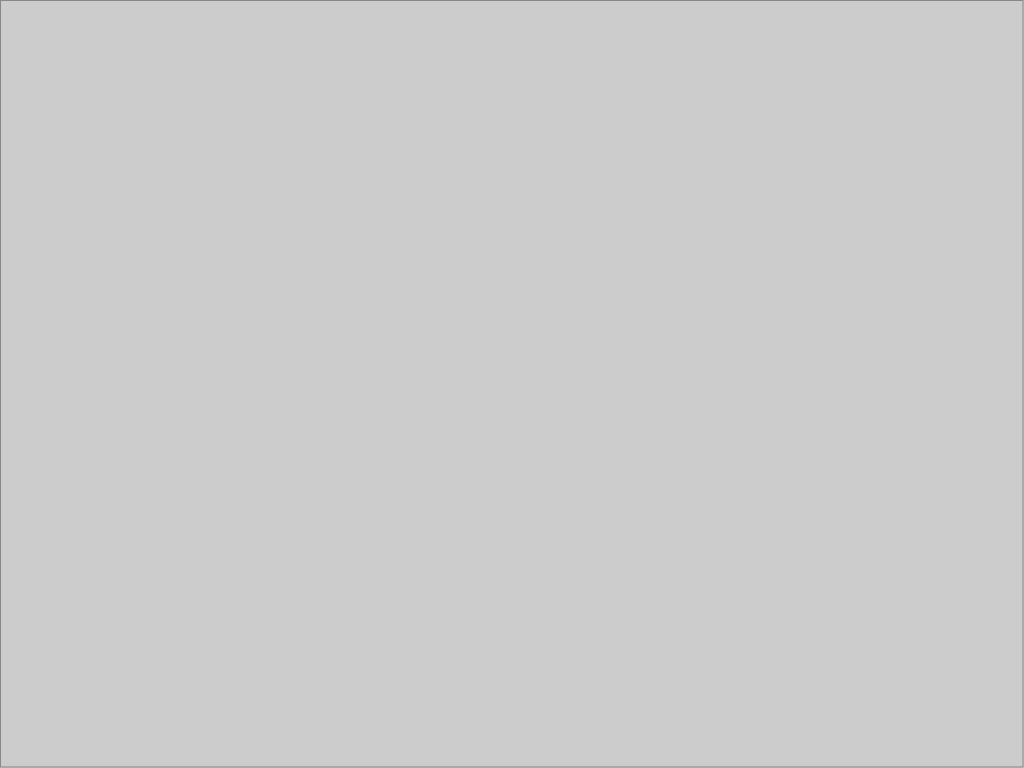
VISUALIZATION Visualization  // 1024x768
    Pie (3360,360 9280x9280)
    Pie (7150,4150 1700x1700)
    Line (8000,8440) (8000,9640)
        p3560616238: MAIN.fbKinematic.X_Visu
        p2738717112: MAIN.fbKinematic.Y_Visu
        p2858320360: MAIN.fbKinematic.Theta_Visu
    Textfield (795,6165 1100x590), "Status :"
    Textfield (775,6825 2840x430), "%s", text variable: GVL_MessageStaus.MessageStaus
    Lamp1 (3935,1815 380x410), style: Lamp-Lamp1-Yellow
END_VISUALIZATION

(* stored: Version 1.1.0.1, ProductVersion 3.1.4024.15
   Visu Visualization: Id {bf080261-e184-4952-90b6-3ab9bf72a664} *)
